Fanuc KAREL source: kd00060.KL

-- PROVISIONAL review KL for V1013-1; original PC SHA256 85b306e1121e9d572326bec6f96117c3b9d167354d8fc59a8972827a10455055
-- Incomplete behavior may be omitted. Consult companion uncertainty JSON. Do not deploy.
PROGRAM KD00060
%NOLOCKGROUP
VAR
  I : INTEGER
  J : INTEGER
  B : BOOLEAN
  R : REAL
  S : STRING[80]
BEGIN
  -- UNRESOLVED_PC offsets 5-18; opcodes 9D,81,18,9D,1B,9D,12,9D,13,04
  -- UNRESOLVED_PC offsets 23-27; opcodes 7F
END KD00060
